(* IEC 61131-3 sources: llm-plc-st-eval/data/calibracion/gemini-3.1-pro-preview/A6/zero_shot, 2 files *)

(* ---- ejec_1.st ---- *)
```iecst
FUNCTION_BLOCK FB_Modos
VAR_INPUT
    selector : INT;
    estadoSeguro : BOOL;
    cmdAuto : ARRAY[0..7] OF BOOL;
    cmdManual : ARRAY[0..7] OF BOOL;
    idxForzado : INT;
    valorForzado : BOOL;
    confirmarForzado : BOOL;
END_VAR

VAR_OUTPUT
    modoActivo : INT :=

(* ---- ejec_3.st ---- *)
```st
FUNCTION_BLOCK FB_Modos
VAR_INPUT
    selector : INT;
    estadoSeguro : BOOL;
    cmdAuto : ARRAY[0..7] OF BOOL;
    cmdManual : ARRAY[0..7] OF BOOL;
    idxForzado : INT;
    valorForzado : BOOL;
    confirmarForzado : BOOL;
END_VAR

VAR_OUTPUT
    modoActivo : INT;
    act
